Fanuc KAREL source: KT00398.KL

PROGRAM KT00398
%NOLOCKGROUP
VAR
  P1: JOINTPOS
  P2: JOINTPOS
  OUT: BOOLEAN
BEGIN
  OUT = P1 <= P2
END KT00398
